(* IEC 61131-3 sources: brew/plant/generated/lite/openplc/plc-packaging, 1 file *)

(* ---- located_vars.st ---- *)
(* Generated by plantgen from plant/plant.yaml (variant lite). Do not edit. *)
(* Analog values are raw registers: engineering value = raw / 10^scaling. *)
(* RIO I/O is at %IX100.0 / %QX100.0 / %IW100 / %QW100 (v3 and v4 alike). *)
(* PLC memory: bits from %QX0.0 (coils), words from %MW0 (holding register qw_count and up, see modbus_slave.json). *)
VAR
  PKG_LINE_PACKML_STATE AT %MW0 : UINT; (* Bottling line PackML state (StateCurrent), None, x1 *)
  PKG_LINE_PACKML_ALM_STATE AT %QX0.0 : BOOL; (* Bottling line PackML state (StateCurrent): state alarm (low) *)
  PKG_LINE_PACKML_MODE AT %MW1 : UINT; (* Bottling line PackML mode (UnitModeCurrent), None, x1 *)
  PKG_LINE_PACKML_CMD AT %MW2 : UINT; (* Bottling line PackML command (CntrlCmd), None, x1 *)
  PKG_LINE_PACKML_MODE_CMD AT %MW3 : UINT; (* Bottling line mode command, None, x1 *)
  PKG_LINE_PACKML_SPEED_SP AT %MW4 : UINT; (* Bottling line speed setpoint (MachSpeed), bottles/min, x10 *)
  PKG_LINE_PACKML_PROCESSED AT %MW5 : UINT; (* Bottles filled this shift (wraps at 65535), None, x1 *)
  PKG_LINE_PACKML_DEFECTIVE AT %MW6 : UINT; (* Bottles rejected this shift (wraps at 65535), None, x1 *)
  PKG_LINE_PACKML_STOP_REASON AT %MW7 : UINT; (* Line stop reason (first-out machine), None, x1 *)
  PKG_LINE_KQ01_OEE AT %MW8 : UINT; (* Shift OEE, %, x10 *)
  PKG_LINE_XS01_RUN AT %QX0.1 : BOOL; (* Line not Stopped or Aborted (alarm suppression) *)
  PKG_FILLER_PACKML_STATE AT %IW100 : UINT; (* Filler PackML state (StateCurrent), None, x1 *)
  PKG_FILLER_PACKML_MODE AT %IW101 : UINT; (* Filler PackML mode (UnitModeCurrent), None, x1 *)
  PKG_FILLER_PACKML_SPEED AT %IW102 : UINT; (* Filler current speed (CurMachSpeed), bottles/min, x10 *)
  PKG_FILLER_PACKML_PROCESSED AT %IW103 : UINT; (* Filler ProdProcessedCount (wraps at 65535), None, x1 *)
  PKG_FILLER_PACKML_DEFECTIVE AT %IW104 : UINT; (* Fill-level inspection rejects (wraps at 65535), None, x1 *)
  PKG_FILLER_PACKML_STOP_REASON AT %IW105 : UINT; (* Filler stop reason (StopReason.ID), None, x1 *)
  PKG_FILLER_PT01_PV AT %IW106 : UINT; (* Filler bowl pressure (absolute), psia, x100 *)
  PKG_FILLER_YA01_PV AT %IX100.0 : BOOL; (* Filler jammed *)
  PKG_FILLER_YA01_ALM_STATE AT %QX0.2 : BOOL; (* Filler jammed: state alarm (low) *)
  PKG_FILLER_LSL01_PV AT %IX100.1 : BOOL; (* Filler bowl low (product supply) *)
  PKG_FILLER_LSL01_ALM_STATE AT %QX0.3 : BOOL; (* Filler bowl low (product supply): state alarm (medium) *)
  PKG_FILLER_XV01_CMD AT %QX100.0 : BOOL; (* Filler product valve (from BBT-202) *)
  PKG_FILLER_PACKML_CMD AT %QW100 : UINT; (* Filler PackML command (CntrlCmd), None, x1 *)
  PKG_FILLER_PACKML_MODE_CMD AT %QW101 : UINT; (* Filler PackML mode command (UnitMode), None, x1 *)
  PKG_FILLER_PACKML_SPEED_SP AT %QW102 : UINT; (* Filler speed setpoint (MachSpeed), bottles/min, x10 *)
  PKG_RINSER_PACKML_STATE AT %IW107 : UINT; (* Rinser PackML state (StateCurrent), None, x1 *)
  PKG_RINSER_PACKML_MODE AT %IW108 : UINT; (* Rinser PackML mode (UnitModeCurrent), None, x1 *)
  PKG_RINSER_PACKML_SPEED AT %IW109 : UINT; (* Rinser current speed (CurMachSpeed), bottles/min, x10 *)
  PKG_RINSER_PACKML_PROCESSED AT %IW110 : UINT; (* Rinser ProdProcessedCount (wraps at 65535), None, x1 *)
  PKG_RINSER_PACKML_DEFECTIVE AT %IW111 : UINT; (* Rinser ProdDefectiveCount (wraps at 65535), None, x1 *)
  PKG_RINSER_PACKML_STOP_REASON AT %IW112 : UINT; (* Rinser stop reason (StopReason.ID), None, x1 *)
  PKG_RINSER_YA01_PV AT %IX100.2 : BOOL; (* Rinser jammed *)
  PKG_RINSER_YA01_ALM_STATE AT %QX0.4 : BOOL; (* Rinser jammed: state alarm (low) *)
  PKG_RINSER_PACKML_CMD AT %QW103 : UINT; (* Rinser PackML command (CntrlCmd), None, x1 *)
  PKG_RINSER_PACKML_MODE_CMD AT %QW104 : UINT; (* Rinser PackML mode command (UnitMode), None, x1 *)
  PKG_RINSER_PACKML_SPEED_SP AT %QW105 : UINT; (* Rinser speed setpoint (MachSpeed), bottles/min, x10 *)
  PKG_CODER_PACKML_STATE AT %IW113 : UINT; (* Date coder PackML state (StateCurrent), None, x1 *)
  PKG_CODER_PACKML_MODE AT %IW114 : UINT; (* Date coder PackML mode (UnitModeCurrent), None, x1 *)
  PKG_CODER_PACKML_SPEED AT %IW115 : UINT; (* Date coder current speed (CurMachSpeed), bottles/min, x10 *)
  PKG_CODER_PACKML_PROCESSED AT %IW116 : UINT; (* Date coder ProdProcessedCount (wraps at 65535), None, x1 *)
  PKG_CODER_PACKML_DEFECTIVE AT %IW117 : UINT; (* Date coder ProdDefectiveCount (wraps at 65535), None, x1 *)
  PKG_CODER_PACKML_STOP_REASON AT %IW118 : UINT; (* Date coder stop reason (StopReason.ID), None, x1 *)
  PKG_CODER_YA01_PV AT %IX100.3 : BOOL; (* Date coder jammed *)
  PKG_CODER_YA01_ALM_STATE AT %QX0.5 : BOOL; (* Date coder jammed: state alarm (low) *)
  PKG_CODER_PACKML_CMD AT %QW106 : UINT; (* Date coder PackML command (CntrlCmd), None, x1 *)
  PKG_CODER_PACKML_MODE_CMD AT %QW107 : UINT; (* Date coder PackML mode command (UnitMode), None, x1 *)
  PKG_CODER_PACKML_SPEED_SP AT %QW108 : UINT; (* Date coder speed setpoint (MachSpeed), bottles/min, x10 *)
  PKG_LABELER_PACKML_STATE AT %IW119 : UINT; (* Labeler PackML state (StateCurrent), None, x1 *)
  PKG_LABELER_PACKML_MODE AT %IW120 : UINT; (* Labeler PackML mode (UnitModeCurrent), None, x1 *)
  PKG_LABELER_PACKML_SPEED AT %IW121 : UINT; (* Labeler current speed (CurMachSpeed), bottles/min, x10 *)
  PKG_LABELER_PACKML_PROCESSED AT %IW122 : UINT; (* Labeler ProdProcessedCount (wraps at 65535), None, x1 *)
  PKG_LABELER_PACKML_DEFECTIVE AT %IW123 : UINT; (* Labeler ProdDefectiveCount (wraps at 65535), None, x1 *)
  PKG_LABELER_PACKML_STOP_REASON AT %IW124 : UINT; (* Labeler stop reason (StopReason.ID), None, x1 *)
  PKG_LABELER_YA01_PV AT %IX100.4 : BOOL; (* Labeler jammed *)
  PKG_LABELER_YA01_ALM_STATE AT %QX0.6 : BOOL; (* Labeler jammed: state alarm (low) *)
  PKG_LABELER_PACKML_CMD AT %QW109 : UINT; (* Labeler PackML command (CntrlCmd), None, x1 *)
  PKG_LABELER_PACKML_MODE_CMD AT %QW110 : UINT; (* Labeler PackML mode command (UnitMode), None, x1 *)
  PKG_LABELER_PACKML_SPEED_SP AT %QW111 : UINT; (* Labeler speed setpoint (MachSpeed), bottles/min, x10 *)
  PKG_PACKER_PACKML_STATE AT %IW125 : UINT; (* Case packer PackML state (StateCurrent), None, x1 *)
  PKG_PACKER_PACKML_MODE AT %IW126 : UINT; (* Case packer PackML mode (UnitModeCurrent), None, x1 *)
  PKG_PACKER_PACKML_SPEED AT %IW127 : UINT; (* Case packer current speed (CurMachSpeed), bottles/min, x10 *)
  PKG_PACKER_PACKML_PROCESSED AT %IW128 : UINT; (* Case packer ProdProcessedCount (wraps at 65535), None, x1 *)
  PKG_PACKER_PACKML_DEFECTIVE AT %IW129 : UINT; (* Case packer ProdDefectiveCount (wraps at 65535), None, x1 *)
  PKG_PACKER_PACKML_STOP_REASON AT %IW130 : UINT; (* Case packer stop reason (StopReason.ID), None, x1 *)
  PKG_PACKER_YA01_PV AT %IX100.5 : BOOL; (* Case packer jammed *)
  PKG_PACKER_YA01_ALM_STATE AT %QX0.7 : BOOL; (* Case packer jammed: state alarm (low) *)
  PKG_PACKER_PACKML_CMD AT %QW112 : UINT; (* Case packer PackML command (CntrlCmd), None, x1 *)
  PKG_PACKER_PACKML_MODE_CMD AT %QW113 : UINT; (* Case packer PackML mode command (UnitMode), None, x1 *)
  PKG_PACKER_PACKML_SPEED_SP AT %QW114 : UINT; (* Case packer speed setpoint (MachSpeed), bottles/min, x10 *)
  PKG_KEG_PACKML_STATE AT %IW131 : UINT; (* Keg washer/filler PackML state (StateCurrent), None, x1 *)
  PKG_KEG_PACKML_MODE AT %IW132 : UINT; (* Keg washer/filler PackML mode (UnitModeCurrent), None, x1 *)
  PKG_KEG_PACKML_PROCESSED AT %IW133 : UINT; (* Kegs filled (wraps at 65535), None, x1 *)
  PKG_KEG_PACKML_DEFECTIVE AT %IW134 : UINT; (* Kegs rejected (wraps at 65535), None, x1 *)
  PKG_KEG_PACKML_STOP_REASON AT %IW135 : UINT; (* Keg washer/filler stop reason, None, x1 *)
  PKG_KEG_TT01_PV AT %IW136 : UINT; (* Keg wash water temperature, degF, x10 *)
  PKG_KEG_YA01_PV AT %IX100.6 : BOOL; (* Keg washer/filler jammed *)
  PKG_KEG_HS01_CMD AT %QX100.1 : BOOL; (* Keg wash heater command *)
  PKG_KEG_PACKML_CMD AT %QW115 : UINT; (* Keg washer/filler PackML command (CntrlCmd), None, x1 *)
  PKG_KEG_PACKML_MODE_CMD AT %QW116 : UINT; (* Keg washer/filler mode command, None, x1 *)
  PKG_CONV_LS01_PV AT %IX100.7 : BOOL; (* Conveyor 1 (depalletizer to rinser) accumulation eye *)
  PKG_CONV_YA01_PV AT %IX101.0 : BOOL; (* Conveyor 1 jam eye *)
  PKG_CONV_HS01_CMD AT %QX100.2 : BOOL; (* Conveyor 1 run command *)
  PKG_CONV_LS02_PV AT %IX101.1 : BOOL; (* Conveyor 2 (filler to coder) accumulation eye *)
  PKG_CONV_YA02_PV AT %IX101.2 : BOOL; (* Conveyor 2 jam eye *)
  PKG_CONV_HS02_CMD AT %QX100.3 : BOOL; (* Conveyor 2 run command *)
  PKG_CONV_LS03_PV AT %IX101.3 : BOOL; (* Conveyor 3 (labeler to packer) accumulation eye *)
  PKG_CONV_YA03_PV AT %IX101.4 : BOOL; (* Conveyor 3 jam eye *)
  PKG_CONV_HS03_CMD AT %QX100.4 : BOOL; (* Conveyor 3 run command *)
  PKG_CONV_LS04_PV AT %IX101.5 : BOOL; (* Conveyor 4 (packer to palletizing) accumulation eye *)
  PKG_CONV_YA04_PV AT %IX101.6 : BOOL; (* Conveyor 4 jam eye *)
  PKG_CONV_HS04_CMD AT %QX100.5 : BOOL; (* Conveyor 4 run command *)
  PKG_PANEL_HS01_PV AT %IW137 : UINT; (* Line command at the operator panel (CntrlCmd while a button is pressed, else 0), None, x1 *)
END_VAR
